// TIA Portal V20 export
// export: Created 2026-10-20T12:45:49.2288816Z, ExportSetting WithDefaults, DisplayName Totally Integrated Automation Portal, DisplayVersion V20 Update 6, DisplayName TIA Portal Openness, DisplayVersion V20 Update 6, DisplayName TIA Portal Version Control Interface, DisplayVersion V20 Update 6, DisplayName SINAMICS Startdrive Advanced, DisplayVersion V20 SP1, DisplayName SINAMICS Startdrive G130, G150, S120, S150, SINAMICS MV, G220, S200, S210, DisplayVersion V20 SP1, DisplayName SINAMICS Startdrive G110M, G120, G120C, G120D, G120P, G115D, DisplayVersion V20 SP1, DisplayName STEP 7 Professional, DisplayVersion V20 Update 6, DisplayName STEP 7 Safety, DisplayVersion V20 Update 2, DisplayName WinCC Basic/Comfort/Advanced, DisplayVersion V20 Update 6, DisplayName WinCC Unified, DisplayVersion V20 Update 6
FUNCTION "PopUp_Screens_2" : Void   // FC63, SCL
{ S7_Optimized_Access := 'TRUE' }
VERSION : 0.1
// stored: AutoNumber true, IsIECCheckEnabled false, SetENOAutomatically false, UDAEnableTagReadback false
   VAR_INPUT
      HMI_No : UInt;
      HMI_Box : UInt;
      Sys_No : UInt;
   END_VAR
BEGIN
   //VTD SETTINGS
   IF "PopUps_DB_1"."VTD_Settings"[#HMI_No].ID <> 0 THEN
       "Settings_DB".VTD_Sys[#Sys_No] := "PopUps_DB_1"."VTD_Settings"[#HMI_No];
       "Settings_Limits_FC"("Settings_DB".VTD_Sys[#Sys_No]);
   END_IF;

   //CONVEYORS SETTINGS
   IF "PopUps_DB_1".ECnv_Settings[#HMI_No].ID <> 0 THEN
       CASE #HMI_Box MOD 10 OF
           1:
               "Settings_DB".LCnv_Sys[#Sys_No].Cnv_Level[1].Cnv1 := "PopUps_DB_1"."Buffer_Cnv_Settings_1"[#HMI_No];
               "Settings_DB".ECnv_Sys[#Sys_No] := "PopUps_DB_1"."ECnv_Settings"[#HMI_No];
               "Settings_DB".LCnv_Sys[#Sys_No].Cnv_Level[1].Cnv2 := "PopUps_DB_1"."Buffer_Cnv_Settings_2"[#HMI_No];
           2:
               "Settings_DB".LCnv_Sys[#Sys_No].Cnv_Level[2].Cnv1 := "PopUps_DB_1"."Buffer_Cnv_Settings_1"[#HMI_No];
               "Settings_DB".ECnv_Sys[#Sys_No] := "PopUps_DB_1"."ECnv_Settings"[#HMI_No];
               "Settings_DB".LCnv_Sys[#Sys_No].Cnv_Level[2].Cnv2 := "PopUps_DB_1"."Buffer_Cnv_Settings_2"[#HMI_No];
           3:
               "Settings_DB".LCnv_Sys[#Sys_No].Cnv_Level[3].Cnv1 := "PopUps_DB_1"."Buffer_Cnv_Settings_1"[#HMI_No];
               "Settings_DB".ECnv_Sys[#Sys_No] := "PopUps_DB_1"."ECnv_Settings"[#HMI_No];
               "Settings_DB".LCnv_Sys[#Sys_No].Cnv_Level[3].Cnv2 := "PopUps_DB_1"."Buffer_Cnv_Settings_2"[#HMI_No];
           4:
               "Settings_DB".LCnv_Sys[#Sys_No].Cnv_Level[4].Cnv1 := "PopUps_DB_1"."Buffer_Cnv_Settings_1"[#HMI_No];
               "Settings_DB".ECnv_Sys[#Sys_No] := "PopUps_DB_1"."ECnv_Settings"[#HMI_No];
               "Settings_DB".LCnv_Sys[#Sys_No].Cnv_Level[4].Cnv2 := "PopUps_DB_1"."Buffer_Cnv_Settings_2"[#HMI_No];
           5:
               "Settings_DB".LCnv_Sys[#Sys_No].Cnv_Level[5].Cnv1 := "PopUps_DB_1"."Buffer_Cnv_Settings_1"[#HMI_No];
               "Settings_DB".ECnv_Sys[#Sys_No] := "PopUps_DB_1"."ECnv_Settings"[#HMI_No];
               "Settings_DB".LCnv_Sys[#Sys_No].Cnv_Level[5].Cnv2 := "PopUps_DB_1"."Buffer_Cnv_Settings_2"[#HMI_No];
           6:
               "Settings_DB".LCnv_Sys[#Sys_No].Cnv_Level[6].Cnv1 := "PopUps_DB_1"."Buffer_Cnv_Settings_1"[#HMI_No];
               "Settings_DB".ECnv_Sys[#Sys_No] := "PopUps_DB_1"."ECnv_Settings"[#HMI_No];
               "Settings_DB".LCnv_Sys[#Sys_No].Cnv_Level[6].Cnv2 := "PopUps_DB_1"."Buffer_Cnv_Settings_2"[#HMI_No];
           7:
               "Settings_DB".LCnv_Sys[#Sys_No].Cnv_Level[7].Cnv1 := "PopUps_DB_1"."Buffer_Cnv_Settings_1"[#HMI_No];
               "Settings_DB".ECnv_Sys[#Sys_No] := "PopUps_DB_1"."ECnv_Settings"[#HMI_No];
               "Settings_DB".LCnv_Sys[#Sys_No].Cnv_Level[7].Cnv2 := "PopUps_DB_1"."Buffer_Cnv_Settings_2"[#HMI_No];
           8:
               "Settings_DB".LCnv_Sys[#Sys_No].Cnv_Level[8].Cnv1 := "PopUps_DB_1"."Buffer_Cnv_Settings_1"[#HMI_No];
               "Settings_DB".ECnv_Sys[#Sys_No] := "PopUps_DB_1"."ECnv_Settings"[#HMI_No];
               "Settings_DB".LCnv_Sys[#Sys_No].Cnv_Level[8].Cnv2 := "PopUps_DB_1"."Buffer_Cnv_Settings_2"[#HMI_No];
       END_CASE;
   END_IF;
END_FUNCTION
